(****************************************************************************************************<br>
© Syntegon Group.<br>
All rights reserved, also regarding any disposal, exploitation, reproduction, editing, distribution,<br>
as well as in the event of applications for industrial property rights.<br>
*****************************************************************************************************<br>
DESCRIPTION:<br>
Parameter set of one Delta robot (ADR 0017): its pose, origin shift, zones, gripper fingers, working area,<br>
limit area and TCP limit area, written by the configurator, taken over when the application allows it.<br>
Typical cycle:<br>
  fb_Delta1Param.m_Register(vio_Manifest := GVL_Config.stManifest, vi_udn_Id := fb_Delta1.m_Id());<br>
  fb_Delta1Param.m_Cycle(vio_Default := Delta1Default, vio_Set := Delta1Set, vi_b_ApplyAllowed := b_Stopped);<br>
  fb_Delta1.m_Configure(vi_lr_BaseRadius := 200, ...);<br>
  fb_Delta1Param.m_PassOn(vio_Visu := fb_Delta1);<br>
The application's pick logic takes its zones from m_Zone / m_Active, not from its own constants.<br>
*****************************************************************************************************<br>
OUTPUT VALUES:<br>
vo_Config is the contract structure the gateway reads and writes at the path in the config manifest.<br>
*****************************************************************************************************<br>
VERSION         ¦ DATE       ¦ NAME      ¦ CHANGE<br>
Syn_Config 1.0.0 ¦ 2026-11-10 ¦ J.Willner ¦ First version<br>
Syn_Config 1.1.0 ¦ 2026-11-10 ¦ J.Willner ¦ m_PassOn, m_Invalid through the shared helpers<br>
Syn_Config 2.0.0 ¦ 2026-11-11 ¦ J.Willner ¦ Gripper fingers with their offsets (ADR 0018)<br>
Syn_Config 2.3.0 ¦ 2026-11-14 ¦ J.Willner ¦ m_Cycle through m_HandleStaging; m_PassOn passes the pose on<br>
****************************************************************************************************)
FUNCTION_BLOCK _FB_ConfigDelta EXTENDS _FB_ConfigComponent
VAR_OUTPUT
	vo_Config							: ST_ConfigDelta;	// contract structure of the gateway
END_VAR

(****************************************************************************************************<br>
© Syntegon Group.<br>
All rights reserved, also regarding any disposal, exploitation, reproduction, editing, distribution,<br>
as well as in the event of applications for industrial property rights.<br>
*****************************************************************************************************<br>
DESCRIPTION:<br>
All effective values (zones, working and limit areas, ...), for the application's own logic.<br>
****************************************************************************************************)
METHOD m_Active : ST_ConfigDeltaParam
m_Active := vo_Config.stActive;
END_METHOD

(****************************************************************************************************<br>
© Syntegon Group.<br>
All rights reserved, also regarding any disposal, exploitation, reproduction, editing, distribution,<br>
as well as in the event of applications for industrial property rights.<br>
*****************************************************************************************************<br>
DESCRIPTION:<br>
A Delta robot.<br>
****************************************************************************************************)
METHOD PROTECTED m_ComponentType : SynVisu.E_VisuComponentType
m_ComponentType := SynVisu.E_VisuComponentType.DELTA;
END_METHOD

(****************************************************************************************************<br>
© Syntegon Group.<br>
All rights reserved, also regarding any disposal, exploitation, reproduction, editing, distribution,<br>
as well as in the event of applications for industrial property rights.<br>
*****************************************************************************************************<br>
DESCRIPTION:<br>
Every cycle: handles a staged set or a reset (a set only while vi_b_ApplyAllowed), keeps the active set in<br>
vio_Set and gives the effective values in vo_Config.stActive: the active set while one is valid, else the<br>
program values vio_Default.<br>
*****************************************************************************************************<br>
OUTPUT VALUES:<br>
TRUE in the cycle a set was taken over or reset.<br>
****************************************************************************************************)
METHOD m_Cycle : BOOL
VAR_IN_OUT CONSTANT
	vio_Default							: ST_ConfigDeltaParam;	// the application's program values
END_VAR
VAR_IN_OUT
	vio_Set								: ST_ConfigDeltaSet;	// the application's VAR PERSISTENT active set
END_VAR
VAR_INPUT
	vi_b_ApplyAllowed					: BOOL;	// [-] a staged set may be taken over now, e.g. while the machine stands
END_VAR
VAR
	b_TempTakeOver						: BOOL;	// the staged set was taken over: copy it
END_VAR
m_Cycle := m_HandleStaging(vio_Staging := vo_Config.stStaging, vio_Status := vo_Config.stStatus, vio_b_Valid := vio_Set.bValid,
	vio_udn_Version := vio_Set.nVersion, vio_udn_LastVersion := vio_Set.nLastVersion, vi_b_ApplyAllowed := vi_b_ApplyAllowed,
	vo_b_TakeOver => b_TempTakeOver);
IF b_TempTakeOver THEN
	vio_Set.stParam := vo_Config.stStaged;
END_IF


(****************************************************************************************************
EFFECTIVE VALUES
****************************************************************************************************)
IF vio_Set.bValid THEN
	vo_Config.stActive := vio_Set.stParam;
ELSE
	vo_Config.stActive := vio_Default;
END_IF
END_METHOD

(****************************************************************************************************<br>
© Syntegon Group.<br>
All rights reserved, also regarding any disposal, exploitation, reproduction, editing, distribution,<br>
as well as in the event of applications for industrial property rights.<br>
*****************************************************************************************************<br>
DESCRIPTION:<br>
Why a staged set cannot be taken over; '' when it can: more zones or fingers than the lists hold, a zone on no<br>
conveyor (id 0), or a finger without a diameter or height.<br>
****************************************************************************************************)
METHOD PROTECTED m_InvalidStaged : STRING(80)
m_InvalidStaged := m_InvalidZones(vio_aZones := vo_Config.stStaged.aZones, vi_un_Count := vo_Config.stStaged.nZoneCount);
IF m_InvalidStaged = '' THEN
	m_InvalidStaged := m_InvalidFingers(vio_aFingers := vo_Config.stStaged.aFingers, vi_un_Count := vo_Config.stStaged.nFingerCount);
END_IF
END_METHOD

(****************************************************************************************************<br>
© Syntegon Group.<br>
All rights reserved, also regarding any disposal, exploitation, reproduction, editing, distribution,<br>
as well as in the event of applications for industrial property rights.<br>
*****************************************************************************************************<br>
DESCRIPTION:<br>
Passes the effective pose, origin shift, working area, limit areas, zones and fingers on to the Delta's<br>
Syn_Visu FB, so the visualisation shows what the machine uses; the arm geometry (hardware) stays with the<br>
application's m_Configure call. Call it after m_Cycle, every cycle; Syn_Visu's config version only changes when a<br>
value does (zones and fingers are cleared only when the set has fewer than the visualisation).<br>
****************************************************************************************************)
METHOD m_PassOn : BOOL
VAR_IN_OUT
	vio_Visu							: SynVisu._FB_VisuDelta;	// the Delta's Syn_Visu FB
END_VAR
m_PassOn := TRUE;
vio_Visu.m_SetPose(vi_Pose := vo_Config.stActive.stPose);
vio_Visu.m_SetOriginShift(vi_lr_X := vo_Config.stActive.stOriginShift.fX, vi_lr_Y := vo_Config.stActive.stOriginShift.fY,
	vi_lr_Z := vo_Config.stActive.stOriginShift.fZ);
vio_Visu.m_SetWorkingArea(vi_lr_Radius := vo_Config.stActive.stWorkingArea.fRadius,
	vi_lr_ZMin := vo_Config.stActive.stWorkingArea.fZMin, vi_lr_ZMax := vo_Config.stActive.stWorkingArea.fZMax,
	vi_lr_ConeHeight := vo_Config.stActive.stWorkingArea.fConeHeight,
	vi_lr_ConeBottomRadius := vo_Config.stActive.stWorkingArea.fConeBottomRadius);
m_PassOnLimitAreas(vio_Visu := vio_Visu, vio_LimitArea := vo_Config.stActive.stLimitArea,
	vio_TcpLimitArea := vo_Config.stActive.stTcpLimitArea);
m_PassOnZones(vio_Visu := vio_Visu, vio_aZones := vo_Config.stActive.aZones, vi_un_Count := vo_Config.stActive.nZoneCount,
	vi_un_VisuCount := vio_Visu.vo_Visu.stConfig.nZoneCount);
m_PassOnFingers(vio_Visu := vio_Visu, vio_aFingers := vo_Config.stActive.aFingers,
	vi_un_Count := vo_Config.stActive.nFingerCount, vi_un_VisuCount := vio_Visu.vo_Visu.stConfig.nFingerCount);
END_METHOD

(****************************************************************************************************<br>
© Syntegon Group.<br>
All rights reserved, also regarding any disposal, exploitation, reproduction, editing, distribution,<br>
as well as in the event of applications for industrial property rights.<br>
*****************************************************************************************************<br>
DESCRIPTION:<br>
Effective pose of the base centre (MCS), for the application's logic.<br>
****************************************************************************************************)
METHOD m_Pose : SynVisu.ST_VisuPose
m_Pose := vo_Config.stActive.stPose;
END_METHOD

(****************************************************************************************************<br>
© Syntegon Group.<br>
All rights reserved, also regarding any disposal, exploitation, reproduction, editing, distribution,<br>
as well as in the event of applications for industrial property rights.<br>
*****************************************************************************************************<br>
DESCRIPTION:<br>
Effective zone vi_un_Zone (1-based, as in Syn_Visu's m_SetZone), for the application's pick and place logic.<br>
*****************************************************************************************************<br>
OUTPUT VALUES:<br>
A zone with nConveyorId = 0 for a number outside 1..m_ZoneCount().<br>
****************************************************************************************************)
METHOD m_Zone : SynVisu.ST_VisuZone
VAR_INPUT
	vi_un_Zone							: UINT;	// [-] 1-based
END_VAR
IF vi_un_Zone >= 1 AND vi_un_Zone <= vo_Config.stActive.nZoneCount
	AND vi_un_Zone <= SynVisu.VISU_GlobalConst_Param.VISU_un_MAX_ZONES
THEN
	m_Zone := vo_Config.stActive.aZones[vi_un_Zone - 1];
END_IF
END_METHOD

(****************************************************************************************************<br>
© Syntegon Group.<br>
All rights reserved, also regarding any disposal, exploitation, reproduction, editing, distribution,<br>
as well as in the event of applications for industrial property rights.<br>
*****************************************************************************************************<br>
DESCRIPTION:<br>
Number of effective zones.<br>
****************************************************************************************************)
METHOD m_ZoneCount : UINT
m_ZoneCount := vo_Config.stActive.nZoneCount;
END_METHOD

END_FUNCTION_BLOCK

(* stored: Version 1.1.0.1
   POU _FB_ConfigDelta: Id {81c755fc-7215-4b2b-96a4-0e696e3e9cd2}, SpecialFunc None
   Method m_Active: Id {892799c0-9099-4e51-ae2c-653fc97e1327}
   Method m_ComponentType: Id {80d968cf-0c4c-48f3-a21c-738e59b951fc}
   Method m_Cycle: Id {55609248-b51c-4028-a529-7706d718eaa7}
   Method m_InvalidStaged: Id {3ba3e387-b7e3-4abe-a51a-555520fb57d1}
   Method m_PassOn: Id {259edc68-b5dc-464d-aec3-df8d64817c9e}
   Method m_Pose: Id {3bfb4653-d713-4059-847e-4083afeb0e49}
   Method m_Zone: Id {0fd56679-9703-4d72-a159-1df3aeda8a30}
   Method m_ZoneCount: Id {433ca3c7-f116-4ad7-90e8-496147f9c07d} *)
